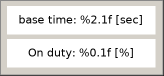
VISUALIZATION vis_FB_DutyCycle_Master  // 164x76
VAR_IN_OUT
	fBaseTime	: REAL;
	fOn_Duty	: REAL;		
END_VAR
    Rectangle (0,0 164x76)
    Textfield (6,5 150x30), "base time: %2.1f [sec]", text variable: fBaseTime
        OnMouseClick: write the text variable via Edit, min 0, max 60
    Textfield (6,38 150x30), "On duty: %0.1f [%]", text variable: fOn_Duty
        OnMouseClick: write the text variable via Edit, min 0, max 100
END_VISUALIZATION

(* stored: Version 1.1.0.1, ProductVersion 3.1.4024.12
   Visu vis_FB_DutyCycle_Master: Id {34165875-6588-4ed4-beb8-484e494e5ade} *)
